Fanuc KAREL source: KT00810.KL

PROGRAM KT00810
%NOLOCKGROUP
VAR
  R1: REAL
  R2: REAL
  OUT: INTEGER
BEGIN
  R1 = 2.0
  R2 = 3.0
  R1 = 2.0
  R2 = 3.0
  OUT = LN(R1)
END KT00810
